(* IEC 61131-3 sources: SortJet_MasterSPS_Aufbau.fbsproj/Device.device.xml.v3^/Plc Logic.plclogic.xml.v3^/Application.application.xml.v3^/09_Station/Shuttle/[101,102] Shuttle/0_Konfig, 7 files *)

(* ---- Antriebsinformationen_Shuttle_101.gvl ---- *)
(* METADATA
{
	"v3Meta": {
		"objectGuid": "b23c52f7-700c-4242-9881-b92df8c5d313"
	}
}
*)
{attribute 'allow_unqualified_access'}
NAMESPACE Antriebsinformationen_Shuttle_101
VAR_GLOBAL

//-------------------------------------------------------------------------------------------------
// ANTRIEBSINFORMATION SHUTTLE
//-------------------------------------------------------------------------------------------------

  apgInfoShuttle101Querfahrt : AntriebsInformationen :=
    (
      wAchsID                                 :=        19,  // Achs ID aus dem EConSet
      stTyp                                   := 'Lateral',  // Typ
      wpSchaltschrank                         :=      3101,  // Daten aus dem Schaltplan
      wpSchaltplanreihe                       :=         2,  // Daten aus dem Schaltplan
      wpSchaltplanseite                       :=        80,  // Daten aus dem Schaltplan
      rpMaxGeschwindigkeit                    :=      3333,  // [mm/s]   Max- Geschwindigkeit für den Automatikbetrieb
      rpHandGeschwindigkeit                   :=       200,  // [mm/s]   Hand- Geschwindigkeit
      rpEinrichtGeschwindigkeit               :=        50,  // [mm/s]   Max Geschwindigkeit während der Einrichtung der Anlage
      rpReferenzGeschwindigkeit               :=        50,  // [mm/s]   Geschwindigkeit für die Referenzfahrt
      rpMaxBeschleunigung                     :=      3000,  // [mm/s^2] Max Beschleunigung
      rpMaxVerzoegerung                       :=      4000,  // [mm/s^2] Max Verzoegerung
      rpMaxRuckzeit                           :=       300,  // [ms]     Ruckzeit des Antriebs
      rpReduzierteBeschleunigung              :=      3500,  // [mm/s^2] Reduzierte Beschleunigung
      rpReduzierteVerzoegerung                :=      4000,  // [mm/s^2] Reduzierte Verzoegerung
      rpGeschwindigkeitMessen                 :=         5,  // [mm/s] Geschwindigkeit beim Scheiben messen
      rpReduzierteGeschwindigkeit             :=       0.0,  // [mm/s]   Reduzierte Geschwindigkeit
      rpBeschleunigungFremdanlage             :=       0.0,  // [mm/s^2] Beschleunigung zu einer Fremdanlage
      rpGeschwindigkeitSystemcheck            :=     500.0,  // [mm/s]   Geschwindigkeit im Systemcheck (nur Glastransport)
      rpGeschwindigkeitSystemcheckReduzierung :=     167.0,  // [mm/s]   Geschwindigkeit im Systemcheck bei belegtem Vorstop-Sensor (nur Glastransport)
      stOptionen                              := ( eEndschalterQuelle    := Endschalterquelle_EN.UMRICHTER, // Hardware-Endschalter: KEINE, UMRICHTER oder SPS
                                                   bVersorgungUeberXVR   := FALSE,                          // XVR-Modus: brueckt Hauptschalter 400 V und LS 230 V
                                                   bBremseLoesenFreigabe := FALSE )                         // Der Antrieb darf über eine Betriebsart die Bremse lösen
    );

  apgInfoShuttle101Glastransport : ARRAY[cWAND_1..cANZAHL_WAENDE] OF AntriebsInformationen := [
    (
      wAchsID                                 :=        20,  // Achs ID aus dem EConSet
      stTyp                                   :=    'Belt',  // Typ
      wpSchaltschrank                         :=      3101,  // Daten aus dem Schaltplan
      wpSchaltplanreihe                       :=         2,  // Daten aus dem Schaltplan
      wpSchaltplanseite                       :=        90,  // Daten aus dem Schaltplan
      rpMaxGeschwindigkeit                    :=      1000,  // [mm/s]   Max- Geschwindigkeit für den Automatikbetrieb
      rpHandGeschwindigkeit                   :=       200,  // [mm/s]   Hand- Geschwindigkeit
      rpReduzierteGeschwindigkeit             :=        67,  // [mm/s]   Reduzierte Geschwindigkeit
      rpReferenzGeschwindigkeit               :=         0,  // [mm/s]   Geschwindigkeit für die Referenzfahrt
      rpEinrichtGeschwindigkeit               :=        50,  // [mm/s]   Max Geschwindigkeit während der Einrichtung der Anlage
      rpMaxBeschleunigung                     :=      1500,  // [mm/s^2] Max Beschleunigung
      rpMaxVerzoegerung                       :=      2000,  // [mm/s^2] Max Verzoegerung
      rpMaxRuckzeit                           :=        50,  // [ms]     Ruckzeit des Antriebs
      rpReduzierteBeschleunigung              :=      1000,  // [mm/s^2] Reduzierte Beschleunigung
      rpReduzierteVerzoegerung                :=      1000,  // [mm/s^2] Reduzierte Verzoegerung
      rpBeschleunigungFremdanlage             :=      1000,  // [mm/s^2] Beschleunigung zu einer Fremdanlage
      rpGeschwindigkeitMessen                 :=       667,  // [mm/s] Geschwindigkeit beim Scheiben messen
      rpGeschwindigkeitSystemcheck            :=     500.0,  // [mm/s]   Geschwindigkeit im Systemcheck (nur Glastransport)
      rpGeschwindigkeitSystemcheckReduzierung :=     167.0,  // [mm/s]   Geschwindigkeit im Systemcheck bei belegtem Vorstop-Sensor (nur Glastransport)
      stOptionen                              := ( eEndschalterQuelle    := Endschalterquelle_EN.KEINE,     // Hardware-Endschalter: KEINE, UMRICHTER oder SPS
                                                   bVersorgungUeberXVR   := FALSE,                          // XVR-Modus: brueckt Hauptschalter 400 V und LS 230 V
                                                   bBremseLoesenFreigabe := FALSE )                         // Der Antrieb darf über eine Betriebsart die Bremse lösen
    )];

  apgInfoShuttle101GlastransportSlave : ARRAY[cWAND_1..cANZAHL_WAENDE] OF AntriebsInformationen := [
    (
      wAchsID                                 :=        65,  // Achs ID aus dem EConSet
      stTyp                                   :=  'BeltSl',  // Typ
      wpSchaltschrank                         :=      3101,  // Daten aus dem Schaltplan
      wpSchaltplanreihe                       :=         2,  // Daten aus dem Schaltplan
      wpSchaltplanseite                       :=        90,  // Daten aus dem Schaltplan
      rpMaxGeschwindigkeit                    :=         0,  // [mm/s]   Max- Geschwindigkeit für den Automatikbetrieb
      rpHandGeschwindigkeit                   :=         0,  // [mm/s]   Hand- Geschwindigkeit
      rpReduzierteGeschwindigkeit             :=         0,  // [mm/s]   Reduzierte Geschwindigkeit
      rpReferenzGeschwindigkeit               :=         0,  // [mm/s]   Geschwindigkeit für die Referenzfahrt
      rpEinrichtGeschwindigkeit               :=         0,  // [mm/s]   Max Geschwindigkeit während der Einrichtung der Anlage
      rpMaxBeschleunigung                     :=         0,  // [mm/s^2] Max Beschleunigung
      rpMaxVerzoegerung                       :=         0,  // [mm/s^2] Max Verzoegerung
      rpMaxRuckzeit                           :=         0,  // [ms]     Ruckzeit des Antriebs
      rpReduzierteBeschleunigung              :=         0,  // [mm/s^2] Reduzierte Beschleunigung
      rpReduzierteVerzoegerung                :=         0,  // [mm/s^2] Reduzierte Verzoegerung
      rpBeschleunigungFremdanlage             :=         0,  // [mm/s^2] Beschleunigung zu einer Fremdanlage
      rpGeschwindigkeitMessen                 :=         0,  // [mm/s] Geschwindigkeit beim Scheiben messen
      rpGeschwindigkeitSystemcheck            :=     500.0,  // [mm/s]   Geschwindigkeit im Systemcheck (nur Glastransport)
      rpGeschwindigkeitSystemcheckReduzierung :=     167.0,  // [mm/s]   Geschwindigkeit im Systemcheck bei belegtem Vorstop-Sensor (nur Glastransport)
      stOptionen                              := ( eEndschalterQuelle    := Endschalterquelle_EN.KEINE,     // Hardware-Endschalter: KEINE, UMRICHTER oder SPS
                                                   bVersorgungUeberXVR   := FALSE,                          // XVR-Modus: brueckt Hauptschalter 400 V und LS 230 V
                                                   bBremseLoesenFreigabe := FALSE )                         // Der Antrieb darf über eine Betriebsart die Bremse lösen
    )];

  apgInfoShuttle101Kippen : AntriebsInformationen :=
    (
      wAchsID                                 :=        65,  // Achs ID aus dem EConSet
      stTyp                                   :=    'Tilt',  // Typ
      wpSchaltschrank                         :=      3101,  // Daten aus dem Schaltplan
      wpSchaltplanreihe                       :=         2,  // Daten aus dem Schaltplan
      wpSchaltplanseite                       :=       110,  // Daten aus dem Schaltplan
      rpMaxGeschwindigkeit                    :=        60,  // [Grad/s]   Max- Geschwindigkeit für den Automatikbetrieb
      rpHandGeschwindigkeit                   :=        60,  // [Grad/s]   Hand- Geschwindigkeit
      rpReduzierteGeschwindigkeit             :=        20,  // [Grad/s]   Reduzierte Geschwindigkeit
      rpEinrichtGeschwindigkeit               :=        20,  // [Grad/s]   Max Geschwindigkeit während der Einrichtung der Anlage
      rpMaxBeschleunigung                     :=        70,  // [Grad/s^2] Max Beschleunigung
      rpMaxVerzoegerung                       :=        70,  // [Grad/s^2] Max Verzoegerung
      rpMaxRuckzeit                           :=       400,  // [ms]     Ruckzeit des Antriebs
      rpReduzierteBeschleunigung              :=        70,  // [Grad/s^2] Reduzierte Beschleunigung
      rpReduzierteVerzoegerung                :=        70,  // [Grad/s^2] Reduzierte Verzoegerung
      rpGeschwindigkeitMessen                 :=         0,  // [Grad/s] Geschwindigkeit beim Scheiben messen
      rpReferenzGeschwindigkeit               :=       0.0,  // [Grad/s]   Geschwindigkeit für die Referenzfahrt
      rpBeschleunigungFremdanlage             :=       0.0,  // [Grad/s^2] Beschleunigung zu einer Fremdanlage
      rpGeschwindigkeitSystemcheck            :=     500.0,  // [mm/s]   Geschwindigkeit im Systemcheck (nur Glastransport)
      rpGeschwindigkeitSystemcheckReduzierung :=     167.0,  // [mm/s]   Geschwindigkeit im Systemcheck bei belegtem Vorstop-Sensor (nur Glastransport)
      stOptionen                              := ( eEndschalterQuelle    := Endschalterquelle_EN.UMRICHTER, // Hardware-Endschalter: KEINE, UMRICHTER oder SPS
                                                   bVersorgungUeberXVR   := FALSE,                          // XVR-Modus: brueckt Hauptschalter 400 V und LS 230 V
                                                   bBremseLoesenFreigabe := FALSE )                         // Der Antrieb darf über eine Betriebsart die Bremse lösen
    );

  apgInfoShuttle101Dickenverstellung : ARRAY[cWAND_1..cANZAHL_WAENDE] OF AntriebsInformationen := [
    (
      wAchsID                                 :=        65,  // Achs ID aus dem EConSet
      stTyp                                   :=    'Wall',  // Typ
      wpSchaltschrank                         :=      3101,  // Daten aus dem Schaltplan
      wpSchaltplanreihe                       :=         2,  // Daten aus dem Schaltplan
      wpSchaltplanseite                       :=       115,  // Daten aus dem Schaltplan
      rpMaxGeschwindigkeit                    :=        60,  // [mm/s]   Max- Geschwindigkeit für den Automatikbetrieb
      rpHandGeschwindigkeit                   :=        60,  // [mm/s]   Hand- Geschwindigkeit
      rpEinrichtGeschwindigkeit               :=        50,  // [mm/s]   Max Geschwindigkeit während der Einrichtung der Anlage
      rpReferenzGeschwindigkeit               :=        50,  // [mm/s]   Geschwindigkeit für die Referenzfahrt
      rpMaxBeschleunigung                     :=       250,  // [mm/s^2] Max Beschleunigung
      rpMaxVerzoegerung                       :=       250,  // [mm/s^2] Max Verzoegerung
      rpMaxRuckzeit                           :=       250,  // [ms]     Ruckzeit des Antriebs
      rpReduzierteBeschleunigung              :=       250,  // [mm/s^2] Reduzierte Beschleunigung
      rpReduzierteVerzoegerung                :=       250,  // [mm/s^2] Reduzierte Verzoegerung
      rpReduzierteGeschwindigkeit             :=       0.0,  // [mm/s]   Reduzierte Geschwindigkeit
      rpBeschleunigungFremdanlage             :=       0.0,  // [mm/s^2] Beschleunigung zu einer Fremdanlage
      rpGeschwindigkeitMessen                 :=       0.0,  // [mm/s] Geschwindigkeit beim Scheiben messen
      rpGeschwindigkeitSystemcheck            :=     500.0,  // [mm/s]   Geschwindigkeit im Systemcheck (nur Glastransport)
      rpGeschwindigkeitSystemcheckReduzierung :=     167.0,  // [mm/s]   Geschwindigkeit im Systemcheck bei belegtem Vorstop-Sensor (nur Glastransport)
      stOptionen                              := ( eEndschalterQuelle    := Endschalterquelle_EN.UMRICHTER, // Hardware-Endschalter: KEINE, UMRICHTER oder SPS
                                                   bVersorgungUeberXVR   := FALSE,                          // XVR-Modus: brueckt Hauptschalter 400 V und LS 230 V
                                                   bBremseLoesenFreigabe := FALSE )                         // Der Antrieb darf über eine Betriebsart die Bremse lösen
    )];

  // Greifer [Ausbaustufe stStationsAufbau.bGreifer]: Achs-ID 65 = nicht vorhanden, Werte aus Schaltplan / Inbetriebnahme eintragen
  apgInfoShuttle101Greifer : ARRAY[cWAND_1..cANZAHL_WAENDE] OF AntriebsInformationen := [
    (
      wAchsID                                 :=        65,  // Achs ID aus dem EConSet
      stTyp                                   := 'Gripper',  // Typ
      wpSchaltschrank                         :=      3101,  // Daten aus dem Schaltplan
      wpSchaltplanreihe                       :=         0,  // Daten aus dem Schaltplan
      wpSchaltplanseite                       :=         0,  // Daten aus dem Schaltplan
      rpMaxGeschwindigkeit                    :=         0,  // [mm/s]   Max- Geschwindigkeit für den Automatikbetrieb
      rpHandGeschwindigkeit                   :=         0,  // [mm/s]   Hand- Geschwindigkeit
      rpReduzierteGeschwindigkeit             :=         0,  // [mm/s]   Reduzierte Geschwindigkeit
      rpReferenzGeschwindigkeit               :=         0,  // [mm/s]   Geschwindigkeit für die Referenzfahrt
      rpEinrichtGeschwindigkeit               :=         0,  // [mm/s]   Max Geschwindigkeit während der Einrichtung der Anlage
      rpMaxBeschleunigung                     :=         0,  // [mm/s^2] Max Beschleunigung
      rpMaxVerzoegerung                       :=         0,  // [mm/s^2] Max Verzoegerung
      rpMaxRuckzeit                           :=         0,  // [ms]     Ruckzeit des Antriebs
      rpReduzierteBeschleunigung              :=         0,  // [mm/s^2] Reduzierte Beschleunigung
      rpReduzierteVerzoegerung                :=         0,  // [mm/s^2] Reduzierte Verzoegerung
      rpBeschleunigungFremdanlage             :=         0,  // [mm/s^2] Beschleunigung zu einer Fremdanlage
      rpGeschwindigkeitMessen                 :=         0,  // [mm/s] Geschwindigkeit beim Scheiben messen
      rpGeschwindigkeitSystemcheck            :=       0.0,  // [mm/s]   Geschwindigkeit im Systemcheck (nur Glastransport)
      rpGeschwindigkeitSystemcheckReduzierung :=       0.0,  // [mm/s]   Geschwindigkeit im Systemcheck bei belegtem Vorstop-Sensor (nur Glastransport)
      stOptionen                              := ( eEndschalterQuelle    := Endschalterquelle_EN.UMRICHTER, // Hardware-Endschalter: KEINE, UMRICHTER oder SPS
                                                   bVersorgungUeberXVR   := FALSE,                          // XVR-Modus: brueckt Hauptschalter 400 V und LS 230 V
                                                   bBremseLoesenFreigabe := FALSE )                         // Der Antrieb darf über eine Betriebsart die Bremse lösen
    )];

END_VAR
END_NAMESPACE

(* ---- Antriebsinformationen_Shuttle_102.gvl ---- *)
(* METADATA
{
	"v3Meta": {
		"objectGuid": "88e35184-05db-4fd2-b301-151a6ca0d672"
	}
}
*)
{attribute 'allow_unqualified_access'}
NAMESPACE Antriebsinformationen_Shuttle_102
VAR_GLOBAL

//-------------------------------------------------------------------------------------------------
// ANTRIEBSINFORMATION SHUTTLE
//-------------------------------------------------------------------------------------------------

  apgInfoShuttle102Querfahrt : AntriebsInformationen :=
    (
      wAchsID                                 :=        21,  // Achs ID aus dem EConSet
      stTyp                                   := 'Lateral',  // Typ
      wpSchaltschrank                         :=      3102,  // Daten aus dem Schaltplan
      wpSchaltplanreihe                       :=         2,  // Daten aus dem Schaltplan
      wpSchaltplanseite                       :=        80,  // Daten aus dem Schaltplan
      rpMaxGeschwindigkeit                    :=      3333,  // [mm/s]   Max- Geschwindigkeit für den Automatikbetrieb
      rpHandGeschwindigkeit                   :=       200,  // [mm/s]   Hand- Geschwindigkeit
      rpEinrichtGeschwindigkeit               :=        50,  // [mm/s]   Max Geschwindigkeit während der Einrichtung der Anlage
      rpReferenzGeschwindigkeit               :=        50,  // [mm/s]   Geschwindigkeit für die Referenzfahrt
      rpMaxBeschleunigung                     :=      3000,  // [mm/s^2] Max Beschleunigung
      rpMaxVerzoegerung                       :=      4000,  // [mm/s^2] Max Verzoegerung
      rpMaxRuckzeit                           :=       300,  // [ms]     Ruckzeit des Antriebs
      rpReduzierteBeschleunigung              :=      3500,  // [mm/s^2] Reduzierte Beschleunigung
      rpReduzierteVerzoegerung                :=      4000,  // [mm/s^2] Reduzierte Verzoegerung
      rpGeschwindigkeitMessen                 :=         5,  // [mm/s] Geschwindigkeit beim Scheiben messen
      rpReduzierteGeschwindigkeit             :=       0.0,  // [mm/s]   Reduzierte Geschwindigkeit
      rpBeschleunigungFremdanlage             :=       0.0,  // [mm/s^2] Beschleunigung zu einer Fremdanlage
      rpGeschwindigkeitSystemcheck            :=     500.0,  // [mm/s]   Geschwindigkeit im Systemcheck (nur Glastransport)
      rpGeschwindigkeitSystemcheckReduzierung :=     167.0,  // [mm/s]   Geschwindigkeit im Systemcheck bei belegtem Vorstop-Sensor (nur Glastransport)
      stOptionen                              := ( eEndschalterQuelle    := Endschalterquelle_EN.UMRICHTER, // Hardware-Endschalter: KEINE, UMRICHTER oder SPS
                                                   bVersorgungUeberXVR   := FALSE,                          // XVR-Modus: brueckt Hauptschalter 400 V und LS 230 V
                                                   bBremseLoesenFreigabe := FALSE )                         // Der Antrieb darf über eine Betriebsart die Bremse lösen
    );

  apgInfoShuttle102Glastransport : ARRAY[cWAND_1..cANZAHL_WAENDE] OF AntriebsInformationen := [
    (
      wAchsID                                 :=        22,  // Achs ID aus dem EConSet
      stTyp                                   :=    'Belt',  // Typ
      wpSchaltschrank                         :=      3102,  // Daten aus dem Schaltplan
      wpSchaltplanreihe                       :=         2,  // Daten aus dem Schaltplan
      wpSchaltplanseite                       :=        90,  // Daten aus dem Schaltplan
      rpMaxGeschwindigkeit                    :=      1000,  // [mm/s]   Max- Geschwindigkeit für den Automatikbetrieb
      rpHandGeschwindigkeit                   :=       200,  // [mm/s]   Hand- Geschwindigkeit
      rpReduzierteGeschwindigkeit             :=        67,  // [mm/s]   Reduzierte Geschwindigkeit
      rpReferenzGeschwindigkeit               :=         0,  // [mm/s]   Geschwindigkeit für die Referenzfahrt
      rpEinrichtGeschwindigkeit               :=        50,  // [mm/s]   Max Geschwindigkeit während der Einrichtung der Anlage
      rpMaxBeschleunigung                     :=      1500,  // [mm/s^2] Max Beschleunigung
      rpMaxVerzoegerung                       :=      2000,  // [mm/s^2] Max Verzoegerung
      rpMaxRuckzeit                           :=        50,  // [ms]     Ruckzeit des Antriebs
      rpReduzierteBeschleunigung              :=      1000,  // [mm/s^2] Reduzierte Beschleunigung
      rpReduzierteVerzoegerung                :=      1000,  // [mm/s^2] Reduzierte Verzoegerung
      rpBeschleunigungFremdanlage             :=      1000,  // [mm/s^2] Beschleunigung zu einer Fremdanlage
      rpGeschwindigkeitMessen                 :=       667,  // [mm/s] Geschwindigkeit beim Scheiben messen
      rpGeschwindigkeitSystemcheck            :=     500.0,  // [mm/s]   Geschwindigkeit im Systemcheck (nur Glastransport)
      rpGeschwindigkeitSystemcheckReduzierung :=     167.0,  // [mm/s]   Geschwindigkeit im Systemcheck bei belegtem Vorstop-Sensor (nur Glastransport)
      stOptionen                              := ( eEndschalterQuelle    := Endschalterquelle_EN.KEINE,     // Hardware-Endschalter: KEINE, UMRICHTER oder SPS
                                                   bVersorgungUeberXVR   := FALSE,                          // XVR-Modus: brueckt Hauptschalter 400 V und LS 230 V
                                                   bBremseLoesenFreigabe := FALSE )                         // Der Antrieb darf über eine Betriebsart die Bremse lösen
    )];

  apgInfoShuttle102GlastransportSlave : ARRAY[cWAND_1..cANZAHL_WAENDE] OF AntriebsInformationen := [
    (
      wAchsID                                 :=        65,  // Achs ID aus dem EConSet
      stTyp                                   :=  'BeltSl',  // Typ
      wpSchaltschrank                         :=      3102,  // Daten aus dem Schaltplan
      wpSchaltplanreihe                       :=         2,  // Daten aus dem Schaltplan
      wpSchaltplanseite                       :=        90,  // Daten aus dem Schaltplan
      rpMaxGeschwindigkeit                    :=         0,  // [mm/s]   Max- Geschwindigkeit für den Automatikbetrieb
      rpHandGeschwindigkeit                   :=         0,  // [mm/s]   Hand- Geschwindigkeit
      rpReduzierteGeschwindigkeit             :=         0,  // [mm/s]   Reduzierte Geschwindigkeit
      rpReferenzGeschwindigkeit               :=         0,  // [mm/s]   Geschwindigkeit für die Referenzfahrt
      rpEinrichtGeschwindigkeit               :=         0,  // [mm/s]   Max Geschwindigkeit während der Einrichtung der Anlage
      rpMaxBeschleunigung                     :=         0,  // [mm/s^2] Max Beschleunigung
      rpMaxVerzoegerung                       :=         0,  // [mm/s^2] Max Verzoegerung
      rpMaxRuckzeit                           :=         0,  // [ms]     Ruckzeit des Antriebs
      rpReduzierteBeschleunigung              :=         0,  // [mm/s^2] Reduzierte Beschleunigung
      rpReduzierteVerzoegerung                :=         0,  // [mm/s^2] Reduzierte Verzoegerung
      rpBeschleunigungFremdanlage             :=         0,  // [mm/s^2] Beschleunigung zu einer Fremdanlage
      rpGeschwindigkeitMessen                 :=         0,  // [mm/s] Geschwindigkeit beim Scheiben messen
      rpGeschwindigkeitSystemcheck            :=     500.0,  // [mm/s]   Geschwindigkeit im Systemcheck (nur Glastransport)
      rpGeschwindigkeitSystemcheckReduzierung :=     167.0,  // [mm/s]   Geschwindigkeit im Systemcheck bei belegtem Vorstop-Sensor (nur Glastransport)
      stOptionen                              := ( eEndschalterQuelle    := Endschalterquelle_EN.KEINE,     // Hardware-Endschalter: KEINE, UMRICHTER oder SPS
                                                   bVersorgungUeberXVR   := FALSE,                          // XVR-Modus: brueckt Hauptschalter 400 V und LS 230 V
                                                   bBremseLoesenFreigabe := FALSE )                         // Der Antrieb darf über eine Betriebsart die Bremse lösen
    )];

  apgInfoShuttle102Kippen : AntriebsInformationen :=
    (
      wAchsID                                 :=        65,  // Achs ID aus dem EConSet
      stTyp                                   :=    'Tilt',  // Typ
      wpSchaltschrank                         :=      3102,  // Daten aus dem Schaltplan
      wpSchaltplanreihe                       :=         2,  // Daten aus dem Schaltplan
      wpSchaltplanseite                       :=       110,  // Daten aus dem Schaltplan
      rpMaxGeschwindigkeit                    :=        60,  // [Grad/s]   Max- Geschwindigkeit für den Automatikbetrieb
      rpHandGeschwindigkeit                   :=        60,  // [Grad/s]   Hand- Geschwindigkeit
      rpReduzierteGeschwindigkeit             :=        20,  // [Grad/s]   Reduzierte Geschwindigkeit
      rpEinrichtGeschwindigkeit               :=        20,  // [Grad/s]   Max Geschwindigkeit während der Einrichtung der Anlage
      rpMaxBeschleunigung                     :=        70,  // [Grad/s^2] Max Beschleunigung
      rpMaxVerzoegerung                       :=        70,  // [Grad/s^2] Max Verzoegerung
      rpMaxRuckzeit                           :=       400,  // [ms]     Ruckzeit des Antriebs
      rpReduzierteBeschleunigung              :=        70,  // [Grad/s^2] Reduzierte Beschleunigung
      rpReduzierteVerzoegerung                :=        70,  // [Grad/s^2] Reduzierte Verzoegerung
      rpGeschwindigkeitMessen                 :=         0,  // [Grad/s] Geschwindigkeit beim Scheiben messen
      rpReferenzGeschwindigkeit               :=       0.0,  // [Grad/s]   Geschwindigkeit für die Referenzfahrt
      rpBeschleunigungFremdanlage             :=       0.0,  // [Grad/s^2] Beschleunigung zu einer Fremdanlage
      rpGeschwindigkeitSystemcheck            :=     500.0,  // [mm/s]   Geschwindigkeit im Systemcheck (nur Glastransport)
      rpGeschwindigkeitSystemcheckReduzierung :=     167.0,  // [mm/s]   Geschwindigkeit im Systemcheck bei belegtem Vorstop-Sensor (nur Glastransport)
      stOptionen                              := ( eEndschalterQuelle    := Endschalterquelle_EN.UMRICHTER, // Hardware-Endschalter: KEINE, UMRICHTER oder SPS
                                                   bVersorgungUeberXVR   := FALSE,                          // XVR-Modus: brueckt Hauptschalter 400 V und LS 230 V
                                                   bBremseLoesenFreigabe := FALSE )                         // Der Antrieb darf über eine Betriebsart die Bremse lösen
    );

  apgInfoShuttle102Dickenverstellung : ARRAY[cWAND_1..cANZAHL_WAENDE] OF AntriebsInformationen := [
    (
      wAchsID                                 :=        65,  // Achs ID aus dem EConSet
      stTyp                                   :=    'Wall',  // Typ
      wpSchaltschrank                         :=      3102,  // Daten aus dem Schaltplan
      wpSchaltplanreihe                       :=         2,  // Daten aus dem Schaltplan
      wpSchaltplanseite                       :=       115,  // Daten aus dem Schaltplan
      rpMaxGeschwindigkeit                    :=        60,  // [mm/s]   Max- Geschwindigkeit für den Automatikbetrieb
      rpHandGeschwindigkeit                   :=        60,  // [mm/s]   Hand- Geschwindigkeit
      rpEinrichtGeschwindigkeit               :=        50,  // [mm/s]   Max Geschwindigkeit während der Einrichtung der Anlage
      rpReferenzGeschwindigkeit               :=        50,  // [mm/s]   Geschwindigkeit für die Referenzfahrt
      rpMaxBeschleunigung                     :=       250,  // [mm/s^2] Max Beschleunigung
      rpMaxVerzoegerung                       :=       250,  // [mm/s^2] Max Verzoegerung
      rpMaxRuckzeit                           :=       250,  // [ms]     Ruckzeit des Antriebs
      rpReduzierteBeschleunigung              :=       250,  // [mm/s^2] Reduzierte Beschleunigung
      rpReduzierteVerzoegerung                :=       250,  // [mm/s^2] Reduzierte Verzoegerung
      rpReduzierteGeschwindigkeit             :=       0.0,  // [mm/s]   Reduzierte Geschwindigkeit
      rpBeschleunigungFremdanlage             :=       0.0,  // [mm/s^2] Beschleunigung zu einer Fremdanlage
      rpGeschwindigkeitMessen                 :=       0.0,  // [mm/s] Geschwindigkeit beim Scheiben messen
      rpGeschwindigkeitSystemcheck            :=     500.0,  // [mm/s]   Geschwindigkeit im Systemcheck (nur Glastransport)
      rpGeschwindigkeitSystemcheckReduzierung :=     167.0,  // [mm/s]   Geschwindigkeit im Systemcheck bei belegtem Vorstop-Sensor (nur Glastransport)
      stOptionen                              := ( eEndschalterQuelle    := Endschalterquelle_EN.UMRICHTER, // Hardware-Endschalter: KEINE, UMRICHTER oder SPS
                                                   bVersorgungUeberXVR   := FALSE,                          // XVR-Modus: brueckt Hauptschalter 400 V und LS 230 V
                                                   bBremseLoesenFreigabe := FALSE )                         // Der Antrieb darf über eine Betriebsart die Bremse lösen
    )];

  // Greifer [Ausbaustufe stStationsAufbau.bGreifer]: zweite Achse des Doppelachsgeraets -90U02
  apgInfoShuttle102Greifer : ARRAY[cWAND_1..cANZAHL_WAENDE] OF AntriebsInformationen := [
    (
      wAchsID                                 :=        23,  // Achs ID aus dem EConSet
      stTyp                                   := 'Gripper',  // Typ
      wpSchaltschrank                         :=      3102,  // Daten aus dem Schaltplan
      wpSchaltplanreihe                       :=         2,  // Daten aus dem Schaltplan
      wpSchaltplanseite                       :=        90,  // Daten aus dem Schaltplan
      rpMaxGeschwindigkeit                    :=      1000,  // [mm/s]   Max- Geschwindigkeit für den Automatikbetrieb
      rpHandGeschwindigkeit                   :=       200,  // [mm/s]   Hand- Geschwindigkeit
      rpReduzierteGeschwindigkeit             :=        67,  // [mm/s]   Reduzierte Geschwindigkeit
      rpReferenzGeschwindigkeit               :=         0,  // [mm/s]   Geschwindigkeit für die Referenzfahrt
      rpEinrichtGeschwindigkeit               :=        50,  // [mm/s]   Max Geschwindigkeit während der Einrichtung der Anlage
      rpMaxBeschleunigung                     :=      1500,  // [mm/s^2] Max Beschleunigung
      rpMaxVerzoegerung                       :=      2000,  // [mm/s^2] Max Verzoegerung
      rpMaxRuckzeit                           :=        50,  // [ms]     Ruckzeit des Antriebs
      rpReduzierteBeschleunigung              :=      1000,  // [mm/s^2] Reduzierte Beschleunigung
      rpReduzierteVerzoegerung                :=      1000,  // [mm/s^2] Reduzierte Verzoegerung
      rpBeschleunigungFremdanlage             :=      1000,  // [mm/s^2] Beschleunigung zu einer Fremdanlage
      rpGeschwindigkeitMessen                 :=       667,  // [mm/s] Geschwindigkeit beim Scheiben messen
      rpGeschwindigkeitSystemcheck            :=     500.0,  // [mm/s]   Geschwindigkeit im Systemcheck (nur Glastransport)
      rpGeschwindigkeitSystemcheckReduzierung :=       0.0,  // [mm/s]   Geschwindigkeit im Systemcheck bei belegtem Vorstop-Sensor (nur Glastransport)
      stOptionen                              := ( eEndschalterQuelle    := Endschalterquelle_EN.UMRICHTER, // Hardware-Endschalter: KEINE, UMRICHTER oder SPS
                                                   bVersorgungUeberXVR   := FALSE,                          // XVR-Modus: brueckt Hauptschalter 400 V und LS 230 V
                                                   bBremseLoesenFreigabe := FALSE )                         // Der Antrieb darf über eine Betriebsart die Bremse lösen
    )];

END_VAR
END_NAMESPACE

(* ---- MK_Shuttle_101.gvl ---- *)
(* METADATA
{
	"v3Meta": {
		"objectGuid": "bf15cf66-58cc-4435-9404-53c8afb203b8"
	}
}
*)
{attribute 'allow_unqualified_access'}
NAMESPACE MK_Shuttle_101
VAR_GLOBAL

//-------------------------------------------------------------------------------------------------
// MASCHINEPARAMETER: SHUTTLE
//-------------------------------------------------------------------------------------------------

  apgMKShuttle101 : Parameter_Station :=
    (
      stStationsNummern                 := ( NummerIntern := 101,                                                                                       // Stationsnummer fuer das MMI und die Stationsangabe der Meldungen
                                             NummerExtern := 1101,                                                                                      // Stationsnummer fuer Bedienermeldungen
                                             NummerSPS    := 101 ),                                                                                     // Stationsnummer SPS-intern (Indizes)
      bDeaktivieren                     := FALSE,                                                                                                       // Station deaktiviert (keine Auftraege, keine Referenzfahrt)
      wMeldungsNummer                   := 600,                                                                                                         // Basis-Meldungsnummer (WatchIO)
      eStationsTyp                      := eInputshuttle,                                                                                               // Typ der Station
      eaAutomatikkreis                  := [eAutomatikkreis_1],                                                                                         // Automatikkreise, zu denen die Station gehoert
      eaSicherheitskreis                := [eSicherheitskreis_1],                                                                                       // Sicherheitskreise, in die die Station eingebunden ist
      // astSicherheitskreisTeilabschaltung
      eSystemcheckZyklus                := eSystemcheckZyklus_1,                                                                                        // In welchem Zyklus des Systemchecks die Station geprueft wird

      stSchnittstellendaten             := (
                                            wVorgaengerStation := cSTATION_DEFAULT,                                                                     // Station vor dieser Station (cSTATION_DYNAMISCH bei mehreren)
                                            wNachfolgerStation := cSTATION_DEFAULT,                                                                     // Station nach dieser Station (cSTATION_DYNAMISCH bei mehreren)
                                            bStationIstShuttle := TRUE                                                                                  // Station ist ein Shuttle
                                          ),

      stStationsOptionen                := (
                                            stSystemcheck := (
                                              bScheibenVermessenSystemCheck           := TRUE,                                                          // Scheiben im Systemcheck vermessen
                                              bScheibeNachSystemcheckAufAuslauf       := TRUE,                                                          // Scheibe nach dem Systemcheck auf den Auslaufsensor fahren
                                              bSystemCheckMitVorgaengerBatchTransport := FALSE,                                                         // derzeit ohne Funktion
                                              bSystemCheckMitNachfolgerBatchTransport := FALSE,                                                         // derzeit ohne Funktion
                                              bOptionSystemCheckScheibeMittigLegen    := FALSE                                                          // derzeit ohne Funktion
                                            ),

                                            // stTransfershuttle
                                            stGlastransport := (
                                              bVortransport                          := FALSE,                                                          // Vortransport aktivieren [Bsp.: Nach einem Eintransport mit gesetztem Bit <Letzte Scheibe>]
                                              bTransportMasterSlaveEintransport      := FALSE,                                                          // derzeit ohne Funktion
                                              bTransportMasterSlaveAustransport      := TRUE,                                                           // Austransport als Slave auf die Achse des Nachfolgers
                                              bGLasUebernahmeSenkrecht               := FALSE,                                                          // RKT - Eintransport in Senkrechter-Position bzw. in Waagerechter- Position [default]
                                              bAustransportISOLinie                  := FALSE,                                                          // Austransport an eine ISO-Linie
                                              bScheibenVermessen                     := FALSE,                                                          // Scheibenmessung am Anlegetisch/Anlegewand
                                              bMessrichtungNegativ                   := FALSE,                                                          // Negative Fahrtrichtung beim Messen
                                              bScheibenmessungEintransport           := FALSE,                                                          // Scheibenmessung beim Eintransport
                                              bScheibenmessungSensorVorabAuslauf     := FALSE                                                           // Scheibenmessung mit SensorVorabAuslauf z.B. Anlegewand
                                            ),

                                            // stAnlegetisch
                                            // stEckuebergabe
                                            // stDrehstation
                                            bVorAbKomponentenAnsteuerung            := TRUE,                                                            // VorAbKomponentenAnsteuerung Auftraege werden bearbeitet
                                            bVerstellungEinAusGefahrenLogikDrehen   := FALSE,                                                           // Verstellung: Logik ein-/ausgefahren gedreht
                                            bLangsamfahrtNockenQuerfahrtAktivieren  := TRUE,                                                            // Querfahrt: Langsamfahrt-Nocken auswerten
                                            bSKBlockierenDurchVorabSensoren         := FALSE,                                                           // Vorab-Sensoren belegt blockieren das Oeffnen des Sicherheitskreises
                                            bStationLeerfahrenBeiSkAnforderung      := FALSE,                                                           // Station bei Anforderung Sicherheitskreis leerfahren
                                            bGlasAbgenommenAutomatischQuittieren    := FALSE,                                                           // derzeit ohne Funktion
                                            bScheibeAbnehmenNachEintransport        := FALSE                                                            // Scheibe nach dem Eintransport wieder abnehmen
                                          ),

      stStationsAufbau                  := (
                                            bGeblase                      := [cANZAHL_WAENDE(TRUE)],                                                    // Ausbaustufe: Geblaese je Wand
                                            bGlastransport                := [cANZAHL_WAENDE(TRUE)],                                                    // Ausbaustufe: Glastransport je Wand
                                            bKippen                       := [cANZAHL_WAENDE(FALSE)],                                                   // Ausbaustufe: Kippen je Wand
                                            bKippenSchuetz                := FALSE,                                                                     // Kippen ueber Schuetz statt Umrichter
                                            bTransportVerstellung         := [cANZAHL_WAENDE(FALSE)],                                                    // Ausbaustufe Shuttle: Transport-/Dickenverstellung je Wand
                                            bWandverstellungMotorisch     := FALSE,                                                                     // Shuttle: Transport-/Wandverstellung mit Antrieb statt pneumatisch
                                            bHub                          := FALSE,                                                                     // Ausbaustufe: Hub der Station
                                            bHubrahmen                    := FALSE,                                                                     // Ausbaustufe: Hubrahmen (Riemen heben/senken)
                                            bDrehen                       := FALSE,                                                                     // Ausbaustufe: Drehen
                                            bQuerachse                    := FALSE,                                                                     // Ausbaustufe: Querachse
                                            bMessachse                    := FALSE,                                                                     // Ausbaustufe: Messachse (Anlegetisch, Anlegewand)
                                            bDruckluft                    := FALSE,                                                                     // Druckluftueberwachung vorhanden
                                            bAnschlag                     := FALSE,                                                                     // Ausbaustufe: Ausrichtanschlaege
                                            bSensorAuslauf                := TRUE,                                                                      // Auslaufsensor vorhanden
                                            bSensorEinlauf                := TRUE,                                                                      // Einlaufsensor vorhanden
                                            bSensorEinlaufStopp           := FALSE,                                                                     // Shuttle: zusaetzlicher Stopp-Sensor am Einlauf (ohne: Einlaufsensor), Gegenstueck zum Auslauf-Stopp im Rueckwaertstransport
                                            bSensorAuslaufStopp           := TRUE,                                                                      // Shuttle: zusaetzlicher Stopp-Sensor am Auslauf (ohne: Auslaufsensor), Verfahrfreigabe und Scheibe hat Shuttle verlassen
                                            bDurchlaufSperreZumNachfolger := FALSE,                                                                     // Ausbaustufe: bewegliche Abschrankung zum Nachfolger
                                            bQuerfahrt                    := TRUE,                                                                      // Ausbaustufe: Querfahrt
                                            bDLSSchmiersystem             := TRUE,                                                                      // Zentralschmierung DLS vorhanden
                                            bGlastransportSlaveVorhanden  := FALSE,                                                                     // Glastransport mit Slave-Antrieb (Meldungen/Ueberwachung Slave)
                                            wHydraulikstation             := 0,                                                                         // Faecherwagen Hydraulik: zugeordnete Hydraulikstation (cHYDRAULIKSTATION_x), 0 = keine
                                            bWandverstellung              := [ FALSE ],                                                                 // Ausbaustufe Station: Wandverstellung je Wand
                                            bRoellchenleiste              := [ FALSE ],                                                                 // Ausbaustufe Station: Roellchenleiste je Wand
                                            bDurchgang                    := FALSE,                                                                     // Station ist Teil eines Durchgangs (belegt = Oeffnen blockiert)
                                            bSlaveAntrieb                 := FALSE,                                                                     // Glastransport mit Slave-Antrieb
                                            bRolltor                      := FALSE,                                                                     // Ausbaustufe Faecherwagen: Rolltor
                                            bKlemmzylinder                := FALSE,                                                                     // Ausbaustufe Faecherwagen: Klemmzylinder fixiert den Oberrahmen beim Ein- und Ausschleusen
                                            bGreifer                      := [cANZAHL_WAENDE(FALSE)],                                                   // Shuttle: Greifer je Wand (Scheibe aus dem Faecherwagen ziehen bzw. hineinschieben)
                                            bRFID                         := FALSE,                                                                     // RFID-Leser vorhanden
                                            bAGV                          := FALSE,                                                                     // Ausbaustufe Faecherwagen: Betrieb mit AGV
                                            bKipparme                     := FALSE,                                                                     // Ausbaustufe: Kipparme
                                            bMessachseAmEndeVomTisch      := FALSE                                                                      // Messachse am Ende des Tisches (Hoehenfehler fragt den Bediener)
                                          ),

      stStationsParameter               := (
                                            rLaengeUebergroesseScheibe              := 5000,                                                            // Shuttle: ab dieser Scheibenlaenge gilt die Scheibe als uebergross [mm]
                                            rMinGlasHoeheAutomatischenEintransport  := 500,                                                             // VSG: Mindesthoehe fuer automatischen Eintransport [mm]
                                            rMinGlasLaengeAutomatischenEintransport := 500,                                                             // VSG: Mindestlaenge fuer automatischen Eintransport [mm]
                                            wMaximaleAnzahlAktiverAuftraege         := 1,                                                               // derzeit ohne Funktion
                                            rMinPosSwEsEingrenzung                  := 0.0,                                                             // Externer zusaetzlicher Software-Endschalter MIN; 0 = inaktiv; darf den MK-MIN nur weiter eingrenzen
                                            rMaxPosSwEsEingrenzung                  := 0.0,                                                             // Externer zusaetzlicher Software-Endschalter MAX; 0 = inaktiv; darf den MK-MAX nur weiter eingrenzen
                                            rPosFreigabePufferAusfahren             := 0.0                                                              // derzeit ohne Funktion
                                          ),

      // stFremdanlage
      stGlasdaten                       := [
                                            (
                                              rlMinGlasLaenge := 350,                                                                                   // minimal zulässige GlasLänge
                                              rlMaxGlasLaenge := 2500,                                                                                  // maximale zulässige GlasLänge
                                              rlMinGlasHoehe  := 190,                                                                                   // minimal zulässige GlasHöhe
                                              rlMaxGlasHoehe  := 1800,                                                                                  // maximale zulässige GlasHöhe
                                              rlMinGlasDicke  := 3,                                                                                   // minimal zulässige GlasDicke
                                              rlMaxGlasDicke  := 12.76,                                                                                    // maximal zulaessige Glasdicke [mm]
                                              rlLaengeMaxGlas := 0.0                                                                                    // maximal zulaessige Glaslaenge [mm]
                                            )],
      // Generische Verfahrfreigabe-Ueberwachung für Shuttle 101:
      astShuttleAnhaltenQuellen             := [
                                                 // [1] Transfershuttle 151 -> Einlaufsensor
                                                 ( bAktiv := TRUE,  wQuellenNummer := cSHUTTLE_151,   wWand := cWAND_1, eSensorTyp := eEinlaufsensor ), // Einlauf- oder Auslaufsensor pruefen
                                                 // [2] Transfershuttle 152 -> Einlaufsensor
                                                 ( bAktiv := TRUE,  wQuellenNummer := cSHUTTLE_152,   wWand := cWAND_1, eSensorTyp := eEinlaufsensor ),
                                                 // [3] Station 202 -> Auslaufsensor
                                                 ( bAktiv := TRUE,  wQuellenNummer := cSTATION_202,   wWand := cWAND_1, eSensorTyp := eAuslaufsensor ),
                                                 // [4] nicht belegt
                                                 ( bAktiv := FALSE ),
                                                 // [5] nicht belegt
                                                 ( bAktiv := FALSE ),
                                                 // [6] nicht belegt
                                                 ( bAktiv := FALSE )
                                               ]
    );

//-------------------------------------------------------------------------------------------------
// SHUTTLE GLASTRANSPORT
//-------------------------------------------------------------------------------------------------

  apgMKShuttle101Glastransport : ARRAY[cWAND_1..cANZAHL_WAENDE] OF Parameter_ShuttleGlastransport := [
    (
      rLaengeStation                    := 2800, // Länge der Station
      rScheibenabstand                  := 300,  // Der Abstand zwischen zwei Scheiben auf der Station
      rWegUeberEinlauf                  := 250,  // Weg ueber den Einlaufsensor hinaus [mm]
      rWegUeberEinlaufRueck             := 50,   // So weit soll ueber den Einlaufsensor gefahren werden
      rUeberwachungEinlaufsensor        := 500,  // Der Abstand vom Auslaufsensor der Vorgängerstation zum Einlaufsensor
      rWegUeberAuslauf                  := 50,   // Weg ueber den Auslaufsensor hinaus [mm]
      rWegUeberAuslaufRueck             := 50,   // So weit soll über den Stopsensore hinaus gefahren werden
      rUeberwachungAuslaufsensor        := 500,  // Beim Vorpositionieren muss der spätestens nach diesem Weg der Auslaufsensor belegt sein
      rWegUeberSensorLetzteScheibe      := 50,   // Weg ueber den Sensor bei der letzten Scheibe [mm]
      rWegUeberSensorSystemCheck        := 15,   // Der Weg der Ueber ein die Sensoren zum vermessen der Scheiben
      rWegUeberwachungSensor            := 500,  // Beschreibt die Wegstrecke die der Ein- Auslaufsensor frei gefahren werden darf bevor ein Fehler gemeldet wird
      rMesstoleranz                     := 5,    // Beschreibt die Strecke ziwischen 2 Sensoren die der Antrieb verfaehrt
      rMessstrecke                      := 2650, // Beschreibt die Strecke ziwischen 2 Sensoren die der Antrieb verfaehrt
      rWegstreckeBisZurVerzoegerung     := 2250  // Beschreibt die Strecke die gefahren werden soll bis der Antrieb abgebremst werden soll
    )];

//-------------------------------------------------------------------------------------------------
// SHUTTLE KIPPEN
//-------------------------------------------------------------------------------------------------

  apgMKShuttle101Kippen : ARRAY[cWAND_1..cANZAHL_WAENDE] OF Parameter_Kippen := [
    (
      tZeitlicheUeberwachungKippen      := TIME#20s0ms, // [ms \ s] Verwendet fuer Antriebe die Ueber einen Schuetz angesteuert werden
      tZeitAntriebsfreigabeErhalten     := TIME#10s0ms, // [ms \ s] Energieeinsparrung: Zeiteinheit nach der die Antriebsfreigabe entzogen werden soll wenn keine Aktion ansteht [1 s = 1000 ms ]
      rToleranz                         := 0.5,         // Toleranz beim Entscheiden der aktuellen Position
      rPosition0Grad                    := 0,           // Waagerechte- Position 0 Grad: Position auf die die Station gehoben werden soll
      rPosition84Grad                   := 0,           // Senkrechte- Position 84 Grad: Position auf die die Station gehoben werden soll
      rPosition88_5Grad                 := 120,         // Senkrechte- Position 84 Grad: Position auf die die Station gehoben werden soll
      rPosition90Grad                   := 178,         // Senkrechte-Position 90 Grad : Position auf die die Station gesenkt werden soll
      rPosition96Grad                   := 0,           // Senkrechte-Position 96 Grad : Position auf die die Station gesenkt werden soll
      bKippenMitSchuetz                 := FALSE        // Kippen per Umrichter oder Schütz
    )];

//-------------------------------------------------------------------------------------------------
// SHUTTLE SCHEIBENFUEHRUNG
//-------------------------------------------------------------------------------------------------

  apgMKShutte101Scheibenfuehrung : ARRAY[cWAND_1..cANZAHL_WAENDE] OF Parameter_Dickenverstellung := [
    (
      rPosition_Minimal                 := 0,   // Position minimal
      rPosition_Mittel                  := 180, // Position mittel
      rPosition_Maximal                 := 180, // Position maximal
      rToleranz                         := 1    // Toleranz beim Positionsvergleich
    )];

//-------------------------------------------------------------------------------------------------
// SHUTTLE GREIFER [Ausbaustufe stStationsAufbau.bGreifer]
//   - Positionen und Wege aus der Inbetriebnahme eintragen (Platzhalter 0)
//   - Aufbau: eine Greiferzange auf der Auslaufseite, Glasrueckhalter nur auf der Greiferseite
//-------------------------------------------------------------------------------------------------

  apgMKShuttle101Greifer : ARRAY[cWAND_1..cANZAHL_WAENDE] OF Parameter_Greifer := [
    (
      eGreiferTyp                                  := eGreiferAuslaufseite, // Greiferseite, wenn der Auftrag keine Seite vorgibt (Systemcheck, Grundstellung)
      tZeitAntriebsfreigabeErhalten                := TIME#10s0ms,          // Energieeinsparung: Zeit nach der die Antriebsfreigabe entzogen wird, wenn keine Aktion ansteht
      tUeberwachungZylinder                        := TIME#5s0ms,           // Zeitueberwachung Greifer aus-/einfahren, Greiferzange und Glasrueckhalter
      tUeberwachungBewegung                        := TIME#60S0MS,          // Zeitueberwachung einer Fahrt der Greiferachse
      tUeberwachungKopplung                        := TIME#10s0ms,          // Zeitueberwachung Kopplung / Entkopplung des Glastransports auf die Greiferachse
      bZangeAbfragenVorhanden                      := FALSE,                // Endlagenabfragen der Greiferzange vorhanden (sonst nur Bewegungszeit)
      tZangeBewegungszeit                          := T#400MS,              // Bewegungszeit der Greiferzange ohne Endlagenabfragen bzw. beim Schliessen auf Glas
      bZangeEinlaufVorhanden                       := FALSE,                // Greiferzange Einlaufseite vorhanden (Ablaeufe ueber die Einlaufseite nur damit)
      bZangeAuslaufVorhanden                       := FALSE,                // Greiferzange Auslaufseite vorhanden (Ablaeufe ueber die Auslaufseite nur damit) - 101 ohne Greifer
      bGlasRueckhalterEinlaufVorhanden             := FALSE,                // Glasrueckhalter Einlaufseite vorhanden (sonst Ausgang aus, gilt als eingefahren)
      bGlasRueckhalterAuslaufVorhanden             := FALSE,                // Glasrueckhalter Auslaufseite vorhanden (sonst Ausgang aus, gilt als eingefahren) - 101 ohne Greifer
      rGrundstellungsPosition_Einlauf              := 0,                    // Grundstellung [Home-Position] Greiferseite Einlauf
      rGrundstellungsPosition_Auslauf              := 0,                    // Grundstellung [Home-Position] Greiferseite Auslauf
      rGrundstellungsPosition_EinlaufEintransport  := 0,                    // Vorabposition vor einem Eintransport ueber die Einlaufseite
      rGrundstellungsPosition_AuslaufEintransport  := 0,                    // Vorabposition vor einem Eintransport ueber die Auslaufseite
      rUebergabePosition_Einlauf                   := 0,                    // Position, bis zu der die Scheibe in den Faecherwagen geschoben wird [Einlaufseite]
      rUebernahmePosition_Einlauf                  := 0,                    // Position, an der die Scheibe im Faecherwagen gegriffen wird [Einlaufseite]
      rUebergabePosition_Auslauf                   := 0,                    // Position, bis zu der die Scheibe in den Faecherwagen geschoben wird [Auslaufseite]
      rUebernahmePosition_Auslauf                  := 0,                    // Position, an der die Scheibe im Faecherwagen gegriffen wird [Auslaufseite]
      rOffsetPosition                              := 0,                    // Abstand der Greiferzange hinter der Glaskante beim Positionieren (Sicherheitsmass gegen Glasbeschaedigung)
      rWegBisZumEinlaufsensor                      := 0,                    // Weg vom Referenzpunkt bis zum Einlaufsensor
      rWegBisZumAuslaufsensor                      := 0,                    // Weg vom Referenzpunkt bis zum Auslaufsensor
      rSicherPositionMinimal                       := 0,                    // Zwischen Minimal und Maximal ragt der Greifer nicht ueber das Shuttle (Querfahrt erlaubt)
      rSicherPositionMaximal                       := 0,                    // Zwischen Minimal und Maximal ragt der Greifer nicht ueber das Shuttle (Querfahrt erlaubt)
      rWegBisZumSicherenEinklappen                 := 0,                    // Weg nach dem Austransport, ab dem der Greifer eingefahren wird [10 - 100 mm]
      rGlasEintransportOffset_Einlauf              := 0,                    // Eintransport letzte Scheibe: Weg ueber den Einlaufsensor [Auftragslaenge + Offset]
      rGlasEintransportOffset_Auslauf              := 0,                    // Eintransport letzte Scheibe: Weg ueber den Auslaufsensor [Auftragslaenge + Offset]
      rGlasEintransportOffset_EinlaufSammeln       := 0,                    // Eintransport weiterer Scheiben: Weg ueber den Einlaufsensor [Auftragslaenge + Offset]
      rGlasEintransportOffset_AuslaufSammeln       := 0,                    // Eintransport weiterer Scheiben: Weg ueber den Auslaufsensor [Auftragslaenge + Offset]
      rLaengeUebergroesseScheibe                   := 0,                    // Ab dieser Scheibenlaenge zieht der Greifer nur bis rPositionUebergrosseScheibe, den Rest zieht der Glastransport
      rPositionUebergrosseScheibe_Einlauf          := 0,                    // Maximale Position mit uebergrosser Scheibe [Einlaufseite]
      rPositionUebergrosseScheibe_Auslauf          := 0,                    // Maximale Position mit uebergrosser Scheibe [Auslaufseite]
      rGreiferAusDemGlasFahrPosition               := 0,                    // Weg, um die geoeffnete Greiferzange vom Glas zu befreien
      rMaximalerWegSensorFreiFahren                := 0,                    // Maximaler Weg der Korrekturfahrt, bis der Sensor frei sein muss
      rWegSensorUeberwachungEintransport           := 0,                    // Nach diesem Weg im Eintransport muss die Scheibe den Sensor belegen, sonst hat der Greifer keine Scheibe
      rKorrekturOffset_Einlauf                     := 0,                    // Weg der Greiferzange in das Glas vor dem Greifen beim Austransport [Einlaufseite]
      rKorrekturOffset_Auslauf                     := 0,                    // Weg der Greiferzange in das Glas vor dem Greifen beim Austransport [Auslaufseite]
      rWegGlasUebergabeposition                    := 0,                    // Weg der Scheibe ueber den Sensor der Greiferseite vor dem Austransport
      rWegGlasUebergabepositionLang                := 0,                    // Wie rWegGlasUebergabeposition, fuer uebergrosse Scheiben
      rLaengeReduzierteGeschwindigkeit             := 0,                    // Austransport: Scheiben ab dieser Laenge komplett mit reduzierter Geschwindigkeit in den Faecherwagen
      rLaengeReduzierteGeschwindigkeitEintransport := 0,                    // Eintransport: Weg mit reduzierter Geschwindigkeit bei schweren Scheiben
      rLaengeReduzierteGeschwindigkeitAustransport := 0,                    // Austransport: erster Weg mit reduzierter Geschwindigkeit in den Faecherwagen
      rMinimalPosition                             := 0,                    // Minimale Zielposition der Greiferachse (Plausibilitaet)
      rMaximalPosition                             := 0                     // Maximale Zielposition der Greiferachse (Plausibilitaet)
    )];

END_VAR
END_NAMESPACE

(* ---- MK_Shuttle_102.gvl ---- *)
(* METADATA
{
	"v3Meta": {
		"objectGuid": "9ea52111-672e-45bd-99aa-d1722119a149"
	}
}
*)
{attribute 'allow_unqualified_access'}
NAMESPACE MK_Shuttle_102
VAR_GLOBAL

//-------------------------------------------------------------------------------------------------
// MASCHINEPARAMETER: SHUTTLE
//-------------------------------------------------------------------------------------------------

  apgMKShuttle102 : Parameter_Station :=
    (
      stStationsNummern                 := ( NummerIntern := 102,                                                                                       // Stationsnummer fuer das MMI und die Stationsangabe der Meldungen
                                             NummerExtern := 1102,                                                                                      // Stationsnummer fuer Bedienermeldungen
                                             NummerSPS    := 102 ),                                                                                     // Stationsnummer SPS-intern (Indizes)
      bDeaktivieren                     := FALSE,                                                                                                        // Station deaktiviert (keine Auftraege, keine Referenzfahrt)
      wMeldungsNummer                   := 650,                                                                                                         // Basis-Meldungsnummer (WatchIO)
      eStationsTyp                      := eOutputshuttle,                                                                                               // Typ der Station
      eaAutomatikkreis                  := [eAutomatikkreis_2],                                                                                         // Automatikkreise, zu denen die Station gehoert
      eaSicherheitskreis                := [eSicherheitskreis_1],                                                                                       // Sicherheitskreise, in die die Station eingebunden ist
      // astSicherheitskreisTeilabschaltung
      eSystemcheckZyklus                := eSystemcheckZyklus_1,                                                                                        // In welchem Zyklus des Systemchecks die Station geprueft wird
      stSchnittstellendaten             := (
                                            wVorgaengerStation := cSTATION_DEFAULT,                                                                     // Station vor dieser Station (cSTATION_DYNAMISCH bei mehreren)
                                            wNachfolgerStation := cSTATION_DEFAULT,                                                                     // Station nach dieser Station (cSTATION_DYNAMISCH bei mehreren)
                                            bStationIstShuttle := TRUE                                                                                  // Station ist ein Shuttle
                                          ),
      stStationsOptionen                := (
                                            stSystemcheck := (
                                              bScheibenVermessenSystemCheck           := TRUE,                                                          // Scheiben im Systemcheck vermessen
                                              bScheibeNachSystemcheckAufAuslauf       := FALSE,                                                         // Scheibe nach dem Systemcheck auf den Auslaufsensor fahren
                                              bSystemCheckMitVorgaengerBatchTransport := FALSE,                                                         // derzeit ohne Funktion
                                              bSystemCheckMitNachfolgerBatchTransport := FALSE,                                                         // derzeit ohne Funktion
                                              bOptionSystemCheckScheibeMittigLegen    := FALSE                                                          // derzeit ohne Funktion
                                            ),
                                            // stTransfershuttle
                                            stGlastransport := (
                                              bVortransport                          := FALSE,                                                          // Vortransport aktivieren [Bsp.: Nach einem Eintransport mit gesetztem Bit <Letzte Scheibe>]
                                              bTransportMasterSlaveEintransport      := FALSE,                                                          // derzeit ohne Funktion
                                              bTransportMasterSlaveAustransport      := FALSE,                                                          // Austransport als Slave auf die Achse des Nachfolgers
                                              bGLasUebernahmeSenkrecht               := FALSE,                                                          // RKT - Eintransport in Senkrechter-Position bzw. in Waagerechter- Position [default]
                                              bAustransportISOLinie                  := FALSE,                                                          // Austransport an eine ISO-Linie
                                              bScheibenVermessen                     := FALSE,                                                          // Scheibenmessung am Anlegetisch/Anlegewand
                                              bMessrichtungNegativ                   := FALSE,                                                          // Negative Fahrtrichtung beim Messen
                                              bScheibenmessungEintransport           := FALSE,                                                          // Scheibenmessung beim Eintransport
                                              bScheibenmessungSensorVorabAuslauf     := FALSE                                                           // Scheibenmessung mit SensorVorabAuslauf z.B. Anlegewand
                                            ),

                                            // stAnlegetisch
                                            // stEckuebergabe
                                            // stDrehstation
                                            bVorAbKomponentenAnsteuerung            := TRUE,                                                            // VorAbKomponentenAnsteuerung Auftraege werden bearbeitet
                                            bVerstellungEinAusGefahrenLogikDrehen   := FALSE,                                                           // Verstellung: Logik ein-/ausgefahren gedreht
                                            bLangsamfahrtNockenQuerfahrtAktivieren  := TRUE,                                                            // Querfahrt: Langsamfahrt-Nocken auswerten
                                            bSKBlockierenDurchVorabSensoren         := FALSE,                                                           // Vorab-Sensoren belegt blockieren das Oeffnen des Sicherheitskreises
                                            bStationLeerfahrenBeiSkAnforderung      := FALSE,                                                           // Station bei Anforderung Sicherheitskreis leerfahren
                                            bGlasAbgenommenAutomatischQuittieren    := FALSE,                                                           // derzeit ohne Funktion
                                            bScheibeAbnehmenNachEintransport        := FALSE                                                            // Scheibe nach dem Eintransport wieder abnehmen
                                          ),
      stStationsAufbau                  := (
                                            bGeblase                      := [cANZAHL_WAENDE(TRUE)],                                                    // Ausbaustufe: Geblaese je Wand
                                            bGlastransport                := [cANZAHL_WAENDE(TRUE)],                                                    // Ausbaustufe: Glastransport je Wand
                                            bKippen                       := [cANZAHL_WAENDE(FALSE)],                                                   // Ausbaustufe: Kippen je Wand
                                            bKippenSchuetz                := FALSE,                                                                     // Kippen ueber Schuetz statt Umrichter
                                            bTransportVerstellung         := [cANZAHL_WAENDE(FALSE)],                                                   // Ausbaustufe Shuttle: Transport-/Dickenverstellung je Wand
                                            bWandverstellungMotorisch     := FALSE,                                                                     // Shuttle: Transport-/Wandverstellung mit Antrieb statt pneumatisch
                                            bHub                          := FALSE,                                                                     // Ausbaustufe: Hub der Station
                                            bHubrahmen                    := FALSE,                                                                     // Ausbaustufe: Hubrahmen (Riemen heben/senken)
                                            bDrehen                       := FALSE,                                                                     // Ausbaustufe: Drehen
                                            bQuerachse                    := FALSE,                                                                     // Ausbaustufe: Querachse
                                            bMessachse                    := FALSE,                                                                     // Ausbaustufe: Messachse (Anlegetisch, Anlegewand)
                                            bDruckluft                    := TRUE,                                                                      // Druckluftueberwachung vorhanden (Druckluft OK %IX114.5)
                                            bAnschlag                     := FALSE,                                                                     // Ausbaustufe: Ausrichtanschlaege
                                            bSensorAuslauf                := TRUE,                                                                      // Auslaufsensor vorhanden
                                            bSensorEinlauf                := TRUE,                                                                      // Einlaufsensor vorhanden
                                            bSensorEinlaufStopp           := FALSE,                                                                     // Shuttle: zusaetzlicher Stopp-Sensor am Einlauf (ohne: Einlaufsensor), Gegenstueck zum Auslauf-Stopp im Rueckwaertstransport
                                            bSensorAuslaufStopp           := TRUE,                                                                      // Shuttle: zusaetzlicher Stopp-Sensor am Auslauf (ohne: Auslaufsensor), Verfahrfreigabe und Scheibe hat Shuttle verlassen
                                            bDurchlaufSperreZumNachfolger := FALSE,                                                                     // Ausbaustufe: bewegliche Abschrankung zum Nachfolger
                                            bQuerfahrt                    := TRUE,                                                                      // Ausbaustufe: Querfahrt
                                            bDLSSchmiersystem             := TRUE,                                                                      // Zentralschmierung DLS vorhanden
                                            bGlastransportSlaveVorhanden  := FALSE,                                                                     // Glastransport mit Slave-Antrieb (Meldungen/Ueberwachung Slave)
                                            wHydraulikstation             := 0,                                                                         // Faecherwagen Hydraulik: zugeordnete Hydraulikstation (cHYDRAULIKSTATION_x), 0 = keine
                                            bWandverstellung              := [ FALSE ],                                                                 // Ausbaustufe Station: Wandverstellung je Wand
                                            bRoellchenleiste              := [ FALSE ],                                                                 // Ausbaustufe Station: Roellchenleiste je Wand
                                            bDurchgang                    := FALSE,                                                                     // Station ist Teil eines Durchgangs (belegt = Oeffnen blockiert)
                                            bSlaveAntrieb                 := FALSE,                                                                     // Glastransport mit Slave-Antrieb
                                            bRolltor                      := FALSE,                                                                     // Ausbaustufe Faecherwagen: Rolltor
                                            bKlemmzylinder                := FALSE,                                                                     // Ausbaustufe Faecherwagen: Klemmzylinder fixiert den Oberrahmen beim Ein- und Ausschleusen
                                            bGreifer                      := [cANZAHL_WAENDE(TRUE)],                                                   // Shuttle: Greifer je Wand (Scheibe aus dem Faecherwagen ziehen bzw. hineinschieben)
                                            bRFID                         := FALSE,                                                                     // RFID-Leser vorhanden
                                            bAGV                          := FALSE,                                                                     // Ausbaustufe Faecherwagen: Betrieb mit AGV
                                            bKipparme                     := FALSE,                                                                     // Ausbaustufe: Kipparme
                                            bMessachseAmEndeVomTisch      := FALSE                                                                      // Messachse am Ende des Tisches (Hoehenfehler fragt den Bediener)
                                          ),
      stStationsParameter               := (
                                            rLaengeUebergroesseScheibe              := 2000,                                                          // Shuttle: ab dieser Scheibenlaenge gilt die Scheibe als uebergross [mm]
                                            rMinGlasHoeheAutomatischenEintransport  := 500,                                                             // VSG: Mindesthoehe fuer automatischen Eintransport [mm]
                                            rMinGlasLaengeAutomatischenEintransport := 500,                                                             // VSG: Mindestlaenge fuer automatischen Eintransport [mm]
                                            wMaximaleAnzahlAktiverAuftraege         := 1,                                                               // derzeit ohne Funktion
                                            rMinPosSwEsEingrenzung                  := 0.0,                                                             // Externer zusaetzlicher Software-Endschalter MIN; 0 = inaktiv; darf den MK-MIN nur weiter eingrenzen
                                            rMaxPosSwEsEingrenzung                  := 0.0,                                                             // Externer zusaetzlicher Software-Endschalter MAX; 0 = inaktiv; darf den MK-MAX nur weiter eingrenzen
                                            rPosFreigabePufferAusfahren             := 0.0                                                              // derzeit ohne Funktion
                                          ),
      // stFremdanlage
      stGlasdaten                       := [
                                            (
                                              rlMinGlasLaenge := 350,                                                                                   // minimal zulässige GlasLänge
                                              rlMaxGlasLaenge := 2500,                                                                                  // maximale zulässige GlasLänge
                                              rlMinGlasHoehe  := 190,                                                                                   // minimal zulässige GlasHöhe
                                              rlMaxGlasHoehe  := 1800,                                                                                  // maximale zulässige GlasHöhe
                                              rlMinGlasDicke  := 3,                                                                                   // minimal zulässige GlasDicke
                                              rlMaxGlasDicke  := 12.76,                                                                                    // maximal zulaessige Glasdicke [mm]
                                              rlLaengeMaxGlas := 0.0                                                                                    // maximal zulaessige Glaslaenge [mm]
                                            )
                                           ],
      // Generische Verfahrfreigabe-Ueberwachung für Shuttle 102:
      astShuttleAnhaltenQuellen             := [
                                                 // [1] Transfershuttle 151 -> Einlaufsensor
                                                 ( bAktiv := TRUE,  wQuellenNummer := cSHUTTLE_151,   wWand := cWAND_1, eSensorTyp := eEinlaufsensor ), // Einlauf- oder Auslaufsensor pruefen
                                                 // [2] Transfershuttle 152 -> Einlaufsensor
                                                 ( bAktiv := TRUE,  wQuellenNummer := cSHUTTLE_152,   wWand := cWAND_1, eSensorTyp := eEinlaufsensor ),
                                                 // [3] Station 202 -> Auslaufsensor
                                                 ( bAktiv := TRUE,  wQuellenNummer := cSTATION_202,   wWand := cWAND_1, eSensorTyp := eAuslaufsensor ),
                                                 // [4] nicht belegt
                                                 ( bAktiv := FALSE ),
                                                 // [5] nicht belegt
                                                 ( bAktiv := FALSE ),
                                                 // [6] nicht belegt
                                                 ( bAktiv := FALSE )
                                               ]
    );

//-------------------------------------------------------------------------------------------------
// SHUTTLE GLASTRANSPORT
//-------------------------------------------------------------------------------------------------

apgMKShuttle102Glastransport : ARRAY[cWAND_1..cANZAHL_WAENDE] OF Parameter_ShuttleGlastransport := [
  (
    rLaengeStation                    := 2800, // Länge der Station
    rScheibenabstand                  := 450,  // Der Abstand zwischen zwei Scheiben auf der Station
    rWegUeberEinlauf                  := 320,  // Weg ueber den Einlaufsensor hinaus [mm]
    rWegUeberEinlaufRueck             := 50,   // So weit soll ueber den Einlaufsensor gefahren werden
    rUeberwachungEinlaufsensor        := 500,  // Der Abstand vom Auslaufsensor der Vorgängerstation zum Einlaufsensor
    rWegUeberAuslauf                  := 50,   // Weg ueber den Auslaufsensor hinaus [mm]
    rWegUeberAuslaufRueck             := 50,   // So weit soll über den Stopsensore hinaus gefahren werden
    rUeberwachungAuslaufsensor        := 500,  // Beim Vorpositionieren muss der spätestens nach diesem Weg der Auslaufsensor belegt sein
    rWegUeberSensorLetzteScheibe      := 50,   // Weg ueber den Sensor bei der letzten Scheibe [mm]
    rWegUeberSensorSystemCheck        := 15,   // Der Weg der Ueber ein die Sensoren zum vermessen der Scheiben
    rWegUeberwachungSensor            := 500,  // Beschreibt die Wegstrecke die der Ein- Auslaufsensor frei gefahren werden darf bevor ein Fehler gemeldet wird
    rMesstoleranz                     := 5,    // Beschreibt die Strecke ziwischen 2 Sensoren die der Antrieb verfaehrt
    rMessstrecke                      := 2750, // Beschreibt die Strecke ziwischen 2 Sensoren die der Antrieb verfaehrt
    rWegstreckeBisZurVerzoegerung     := 2250  // Beschreibt die Strecke die gefahren werden soll bis der Antrieb abgebremst werden soll
  )];

//-------------------------------------------------------------------------------------------------
// SHUTTLE KIPPEN
//-------------------------------------------------------------------------------------------------

apgMKShuttle102Kippen : ARRAY[cWAND_1..cANZAHL_WAENDE] OF Parameter_Kippen := [
  (
    tZeitlicheUeberwachungKippen      := TIME#20s0ms, // [ms \ s] Verwendet fuer Antriebe die Ueber einen Schuetz angesteuert werden
    tZeitAntriebsfreigabeErhalten     := TIME#10s0ms, // [ms \ s] Energieeinsparrung: Zeiteinheit nach der die Antriebsfreigabe entzogen werden soll wenn keine Aktion ansteht [1 s = 1000 ms ]
    rToleranz                         := 0.5,         // Toleranz beim Entscheiden der aktuellen Position
    rPosition0Grad                    := 0,           // Waagerechte- Position 0 Grad: Position auf die die Station gehoben werden soll
    rPosition84Grad                   := 0,           // Senkrechte- Position 84 Grad: Position auf die die Station gehoben werden soll
    rPosition88_5Grad                 := 120,         // Senkrechte- Position 84 Grad: Position auf die die Station gehoben werden soll
    rPosition90Grad                   := 178,         // Senkrechte-Position 90 Grad : Position auf die die Station gesenkt werden soll
    rPosition96Grad                   := 0,           // Senkrechte-Position 96 Grad : Position auf die die Station gesenkt werden soll
    bKippenMitSchuetz                 := FALSE        // Kippen per Umrichter oder Schütz
  )];
//-------------------------------------------------------------------------------------------------
// SHUTTLE SCHEIBENFUEHRUNG
//-------------------------------------------------------------------------------------------------

  apgMKShutte102Scheibenfuehrung : ARRAY[cWAND_1..cANZAHL_WAENDE] OF Parameter_Dickenverstellung := [
    (
      rPosition_Minimal                 := 0,   // Position minimal
      rPosition_Mittel                  := 180, // Position mittel
      rPosition_Maximal                 := 180, // Position maximal
      rToleranz                         := 1    // Toleranz beim Positionsvergleich
    )];

//-------------------------------------------------------------------------------------------------
// SHUTTLE GREIFER [Ausbaustufe stStationsAufbau.bGreifer]
//   - Positionen und Wege aus der Inbetriebnahme eintragen (Platzhalter 0)
//   - Aufbau: eine Greiferzange auf der Auslaufseite, Glasrueckhalter nur auf der Greiferseite
//-------------------------------------------------------------------------------------------------

  apgMKShuttle102Greifer : ARRAY[cWAND_1..cANZAHL_WAENDE] OF Parameter_Greifer := [
    (
      eGreiferTyp                                  := eGreiferAuslaufseite, // Greiferseite, wenn der Auftrag keine Seite vorgibt (Systemcheck, Grundstellung)
      tZeitAntriebsfreigabeErhalten                := TIME#180S,            // Energieeinsparung: Zeit nach der die Antriebsfreigabe entzogen wird, wenn keine Aktion ansteht
      tUeberwachungZylinder                        := TIME#5s0ms,           // Zeitueberwachung Greifer aus-/einfahren, Greiferzange und Glasrueckhalter
      tUeberwachungBewegung                        := TIME#60s0ms,          // Zeitueberwachung einer Fahrt der Greiferachse
      tUeberwachungKopplung                        := TIME#10s0ms,          // Zeitueberwachung Kopplung / Entkopplung des Glastransports auf die Greiferachse
      bZangeAbfragenVorhanden                      := FALSE,                // Endlagenabfragen der Greiferzange vorhanden (sonst nur Bewegungszeit)
      tZangeBewegungszeit                          := T#400MS,              // Bewegungszeit der Greiferzange ohne Endlagenabfragen bzw. beim Schliessen auf Glas
      bZangeEinlaufVorhanden                       := FALSE,                // Greiferzange Einlaufseite vorhanden (Ablaeufe ueber die Einlaufseite nur damit)
      bZangeAuslaufVorhanden                       :=  TRUE,                // Greiferzange Auslaufseite vorhanden (Ablaeufe ueber die Auslaufseite nur damit)
      bGlasRueckhalterEinlaufVorhanden             := FALSE,                // Glasrueckhalter Einlaufseite vorhanden (sonst Ausgang aus, gilt als eingefahren)
      bGlasRueckhalterAuslaufVorhanden             :=  TRUE,                // Glasrueckhalter Auslaufseite vorhanden (sonst Ausgang aus, gilt als eingefahren)
      rGrundstellungsPosition_Einlauf              :=    25,                // Grundstellung [Home-Position] Greiferseite Einlauf
      rGrundstellungsPosition_Auslauf              :=  1780,                // Grundstellung [Home-Position] Greiferseite Auslauf
      rGrundstellungsPosition_EinlaufEintransport  :=    25,                // Vorabposition vor einem Eintransport ueber die Einlaufseite
      rGrundstellungsPosition_AuslaufEintransport  :=  1780,                // Vorabposition vor einem Eintransport ueber die Auslaufseite
      rUebergabePosition_Einlauf                   :=    25,                // Position, bis zu der die Scheibe in den Faecherwagen geschoben wird [Einlaufseite]
      rUebernahmePosition_Einlauf                  :=    25,                // Position, an der die Scheibe im Faecherwagen gegriffen wird [Einlaufseite]
      rUebergabePosition_Auslauf                   :=  2350,                // Position, bis zu der die Scheibe in den Faecherwagen geschoben wird [Auslaufseite]
      rUebernahmePosition_Auslauf                  :=  2350,                // Position, an der die Scheibe im Faecherwagen gegriffen wird [Auslaufseite]
      rOffsetPosition                              :=    15,                // Abstand der Greiferzange hinter der Glaskante beim Positionieren (Sicherheitsmass gegen Glasbeschaedigung)
      rWegBisZumEinlaufsensor                      :=    25,                // Weg vom Referenzpunkt bis zum Einlaufsensor
      rWegBisZumAuslaufsensor                      :=  2075,                // Weg vom Referenzpunkt bis zum Auslaufsensor
      rSicherPositionMinimal                       :=    25,                // Zwischen Minimal und Maximal ragt der Greifer nicht ueber das Shuttle (Querfahrt erlaubt)
      rSicherPositionMaximal                       :=  2195,                // Zwischen Minimal und Maximal ragt der Greifer nicht ueber das Shuttle (Querfahrt erlaubt)
      rWegBisZumSicherenEinklappen                 :=    50,                // Weg nach dem Austransport, ab dem der Greifer eingefahren wird [10 - 100 mm]
      rGlasEintransportOffset_Einlauf              :=    50,                // Eintransport letzte Scheibe: Weg ueber den Einlaufsensor [Auftragslaenge + Offset]
      rGlasEintransportOffset_Auslauf              :=    50,                // Eintransport letzte Scheibe: Weg ueber den Auslaufsensor [Auftragslaenge + Offset]
      rGlasEintransportOffset_EinlaufSammeln       :=   450,                // Eintransport weiterer Scheiben: Weg ueber den Einlaufsensor [Auftragslaenge + Offset]
      rGlasEintransportOffset_AuslaufSammeln       :=   370,                // Eintransport weiterer Scheiben: Weg ueber den Auslaufsensor [Auftragslaenge + Offset]
      rLaengeUebergroesseScheibe                   :=  2000,              // Ab dieser Scheibenlaenge zieht der Greifer nur bis rPositionUebergrosseScheibe, den Rest zieht der Glastransport
      rPositionUebergrosseScheibe_Einlauf          :=   500,                // Maximale Position mit uebergrosser Scheibe [Einlaufseite]
      rPositionUebergrosseScheibe_Auslauf          :=   500,                // Maximale Position mit uebergrosser Scheibe [Auslaufseite]
      rGreiferAusDemGlasFahrPosition               :=    50,                // Weg, um die geoeffnete Greiferzange vom Glas zu befreien
      rMaximalerWegSensorFreiFahren                :=   200,                // Maximaler Weg der Korrekturfahrt, bis der Sensor frei sein muss
      rWegSensorUeberwachungEintransport           :=   300,                // Nach diesem Weg im Eintransport muss die Scheibe den Sensor belegen, sonst hat der Greifer keine Scheibe
      rKorrekturOffset_Einlauf                     :=    10,                // Weg der Greiferzange in das Glas vor dem Greifen beim Austransport [Einlaufseite]
      rKorrekturOffset_Auslauf                     :=    10,                // Weg der Greiferzange in das Glas vor dem Greifen beim Austransport [Auslaufseite]
      rWegGlasUebergabeposition                    :=    50,                // Weg der Scheibe ueber den Sensor der Greiferseite vor dem Austransport
      rWegGlasUebergabepositionLang                :=   500,                // Wie rWegGlasUebergabeposition, fuer uebergrosse Scheiben
      rLaengeReduzierteGeschwindigkeit             :=  2000,                // Austransport: Scheiben ab dieser Laenge komplett mit reduzierter Geschwindigkeit in den Faecherwagen
      rLaengeReduzierteGeschwindigkeitEintransport :=   300,                // Eintransport: Weg mit reduzierter Geschwindigkeit bei schweren Scheiben
      rLaengeReduzierteGeschwindigkeitAustransport :=   300,                // Austransport: erster Weg mit reduzierter Geschwindigkeit in den Faecherwagen
      rMinimalPosition                             :=    25,                // Minimale Zielposition der Greiferachse (Plausibilitaet)
      rMaximalPosition                             :=  2390                 // Maximale Zielposition der Greiferachse (Plausibilitaet)
    )];

END_VAR
END_NAMESPACE
